FUNCTION_BLOCK FsWrite (* Write a byte array as file to the file server *)
  (* Standard: 61499-2; Description: Uses iso_FscWriteFileToServer() or iso_FscAppendFileToServer() of the CCI ISOBUS driver (ISO 11783-13). \n Client is NmDestin.s16OwnCfHnd, file server is NmDestin.s16Handle (e.g. found with NmGetCfInfo, NAME function 61). \n The connection is opened and closed by the driver. One job at a time: REQ during a job gives ERR with s16Status E_BUSY. \n Every REQ ends with exactly one CNF or ERR. \n The first u32Length bytes of Data are written. *)
  (* Version 1.0, 2026-11-25, Franz Höpfinger, initial API and implementation and/or initial documentation *)
  PACKAGE isobus::fs;
  IMPORT isobus::pgn::ISONETEVENT_T;
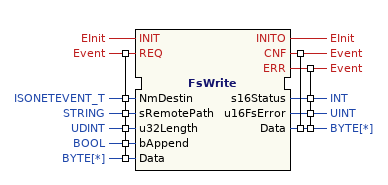
  EVENT_INPUT
    INIT : EInit; (* Service Initialization *)
    REQ WITH NmDestin, sRemotePath, u32Length, bAppend, Data; (* Write the file *)
  END_EVENT
  EVENT_OUTPUT
    INITO : EInit; (* Initialization Confirm *)
    CNF WITH Data; (* File written *)
    ERR WITH s16Status, u16FsError, Data; (* Job failed *)
  END_EVENT
  VAR_INPUT
    NmDestin : isobus::pgn::ISONETEVENT_T; (* Client (s16OwnCfHnd) and file server (s16Handle) *)
    sRemotePath : STRING; (* Path on the file server, e.g. \\USB\data\a.csv *)
    u32Length : UDINT; (* Number of bytes of Data to write *)
    bAppend : BOOL; (* FALSE: replace the file, TRUE: append *)
  END_VAR
  VAR_OUTPUT
    s16Status : INT; (* With ERR: driver return value or own error (E_BUSY, E_RANGE, E_OVERFLOW) *)
    u16FsError : UINT; (* With ERR: file server or client error (ISO 11783-13 B.9, 6400 ff. client) *)
  END_VAR
  VAR_IN_OUT
    Data : ARRAY [*] OF BYTE; (* File content *)
  END_VAR
END_FUNCTION_BLOCK
